FUNCTION_BLOCK FB_Buffer2_4 IMPLEMENTS ITF_Buffer2_4
VAR_INPUT
END_VAR
VAR_OUTPUT
END_VAR
VAR
END_VAR

{warning 'Add method implementation '}
METHOD Aborted : BOOL
END_METHOD

{warning 'Add method implementation '}
METHOD Aborting : BOOL
END_METHOD

{warning 'Add method implementation '}
METHOD Clearing : BOOL
END_METHOD

{warning 'Add method implementation '}
METHOD Execute : BOOL
END_METHOD

{warning 'Add method implementation '}
METHOD Held : BOOL
END_METHOD

{warning 'Add method implementation '}
METHOD Holding : BOOL
END_METHOD

{warning 'Add method implementation '}
METHOD Idle : BOOL
END_METHOD

{warning 'Add method implementation '}
METHOD Resetting : BOOL
END_METHOD

{warning 'Add method implementation '}
METHOD Starting : BOOL
END_METHOD

{warning 'Add method implementation '}
METHOD Stopped : BOOL
END_METHOD

{warning 'Add method implementation '}
METHOD Stopping : BOOL
END_METHOD

{warning 'Add method implementation '}
METHOD Suspended : BOOL
END_METHOD

{warning 'Add method implementation '}
METHOD Suspending : BOOL
END_METHOD

{warning 'Add method implementation '}
METHOD Unholding : BOOL
END_METHOD

{warning 'Add method implementation '}
METHOD Unsuspending : BOOL
END_METHOD

END_FUNCTION_BLOCK

(* stored: Version 1.1.0.1
   POU FB_Buffer2_4: Id {85233061-3399-48bc-adeb-5452bf49870d}, SpecialFunc None
   Folder Methods: Id {2a6015b8-08d0-4b03-aeea-006f8f194aff}
   Method Aborted: Id {2ebeca73-8fac-456a-a7ed-e89a58580cd9}
   Method Aborting: Id {4e4319a7-70b5-43db-8141-c749dfd36c1d}
   Method Clearing: Id {cc4d4c18-f8bf-438a-b70b-6ea20efc7ccf}
   Method Execute: Id {064eaf4d-547c-48e9-a1c7-ebcf1d12dca1}
   Method Held: Id {2ddeec7f-95b5-44f9-b76b-458fe7ece936}
   Method Holding: Id {21c36e0a-c9f6-474a-940c-7ff1bae2f1c6}
   Method Idle: Id {13e96ba2-3274-48cb-9d8d-25e40a7916ea}
   Method Resetting: Id {b55c70df-ecef-44b0-a694-7d16d9e19634}
   Method Starting: Id {bc7fe667-1bb1-490d-8a62-571071c06e76}
   Method Stopped: Id {2380e4c8-6423-4d1b-8020-9ff959cc1734}
   Method Stopping: Id {2cff1f0e-34d6-4e24-9505-5e88ec77a62e}
   Method Suspended: Id {cbf60056-93b2-478a-8f59-89146df3ba88}
   Method Suspending: Id {9028c479-6e8b-4f02-ad2a-9becab1a6e72}
   Method Unholding: Id {e4d7ad9d-2b7f-49f3-8b14-5964a839d612}
   Method Unsuspending: Id {eacaf4c7-df15-4648-80cc-8afc8810550f} *)
